Fanuc KAREL source: KA00070.KL

PROGRAM KA00070
%NOLOCKGROUP
VAR
  SRC: XYZWPR
  DST: CONFIG
BEGIN
  SRC.X = 1.0
  DST = SRC
END KA00070
